// TIA Portal V19 export
// export: Created 2000-01-01T00:00:00.0000000Z, ExportSetting None
FUNCTION "FC_Rung" : Void   // FC42, LAD
{ S7_Optimized_Access := 'TRUE' }
   VAR_INPUT
      Local : Int;
   END_VAR
   VAR_TEMP   // added for the SCL form of the ladder/FBD networks
      _w1 : Bool;
   END_VAR
BEGIN

REGION Network 1
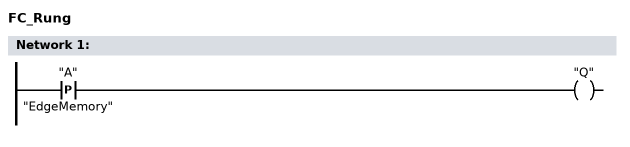
   #_w1 := "A" AND NOT "EdgeMemory";   // rising edge of "A"
   "EdgeMemory" := "A";
   "Q" := #_w1;
END_REGION
END_FUNCTION
